VISUALIZATION FP_Conveyor  // 2x2
END_VISUALIZATION

(* stored: Version 1.1.0.1
   Visu FP_Conveyor: Id {a996403e-7bae-44dc-b93b-b0426081b2c4} *)
